Universal Robots URScript: T013_deepseek-coder-v2_16b_baseline_rep1.urscript

# Define the sequence of moves for the task
def move_joint():
    motion_group.movej([0, -pi/4, pi/3, -pi/4, pi/2, 0], 200, 1.5, avoid_singular=True)

def move_linear(pose):
    motion_group.movel(pose, 220, 1.5, relative=False, avoid_singular=True)

# Define the poses for each move in sequence
home_pose = [0, -pi/4, pi/3, -pi/4, pi/2, 0]
above_staging_pose = [0.2, 0.1, 0.2, 0, 0, 0]
descend_to_pick_pose = [0.2, 0.1, 0.1, 0, 0, 0]
lift_pose = [0.2, 0.1, 0.3, 0, 0, 0]
transit_to_pallet_pose = [0.4, -0.2, 0.3, 0, 0, 0]
# Add more poses as needed...

# Define the safety zone (confinement) if required
safety_zone(0.1)

# Execute the sequence of moves
move_joint()
move_linear(above_staging_pose)
move_linear(descend_to_pick_pose)
move_linear(lift_pose)
move_linear(transit_to_pallet_pose)
# Add more move_linear calls for subsequent poses...
